// TIA Portal V15.1 export
// export: Created 2026-09-17T17:40:11.5857197Z, ExportSetting WithDefaults, DisplayName Totally Integrated Automation Portal, DisplayVersion V15.1, DisplayName TIA Portal Openness, DisplayVersion V15.1, DisplayName STEP 7 Professional, DisplayVersion V15.1, DisplayName WinCC Professional, DisplayVersion V15.1
Screen "faults"  1024x768, Number=5
  ScreenLayer 
    Button "Button_1" at 31,675 size 90x44  Mode=Text, StyleItem=Button, TextOff="End RT", TextOn="Text"
      on Press: StopRuntime(Mode := 0)
    Button "Button_2" at 31,619 size 90x44  Mode=Text, StyleItem=Button, TextOff="Back", TextOn="Text"
      on Press: ActivateScreen(Screen name := Start Screen, Object number := 0)
